SUBAPPLICATION Softkey_Aux_IXA_TO_DataPanel_QXA_BG (* SoftKey ODER AUX auf DataPanel-MI-Ausgang, Hintergrundfarbe SoftKey+AUX Gruen/Weiss, 2 AX-Ausgaenge *)
  (* Standard: 61499-2; Description: Copyright (c) 2026 Meisterschulen am Ostbahnhof This program and the accompanying materials are made available under the terms of the Eclipse Public License 2.0 which is available at https://www.eclipse.org/legal/epl-2.0/ SPDX-License-Identifier: EPL-2.0 *)
  (* Version 1.0, 2026-10-31, Franz Höpfinger, Meisterschulen am Ostbahnhof, Aus Getreidehacke func/Manual/ManFuncTast2 in MyLib::sys verschoben und umbenannt, INIT/INITO/QI/QO ergaenzt, Output und u8SAMember als Parameter. *)
  PACKAGE MyLib::sys;
  IMPORT isobus::UT::Q::const::IDs::ID_NULL;
  IMPORT DataPanel::io::MI::DQ::DataPanel_MI_DO_S;
  IMPORT DataPanel::io::MI::DQ::DataPanel_MI_DO;
  IMPORT DataPanel::io::MI::const::MI;
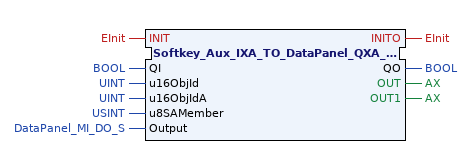
  EVENT_INPUT
    INIT : EInit; (* Initialization Request *)
  END_EVENT
  EVENT_OUTPUT
    INITO : EInit; (* Initialization Confirm *)
  END_EVENT
  VAR_INPUT
    QI : BOOL := TRUE; (* Quality Input - TRUE to enable service *)
    u16ObjId : UINT := ID_NULL; (* Object ID SoftKey *)
    u16ObjIdA : UINT := ID_NULL; (* Object ID AuxFunction2 *)
    u8SAMember : USINT := MI::MI_00; (* DataPanel-MI-Modul (Source Address) *)
    Output : DataPanel::io::MI::DQ::DataPanel_MI_DO_S := DataPanel_MI_DO::Invalid; (* DataPanel-MI-Ausgang *)
  END_VAR
  VAR_OUTPUT
    QO : BOOL; (* Quality Output - TRUE if service executed successfully *)
  END_VAR
  PLUGS
    OUT : adapter::types::unidirectional::AX; (* SoftKey ODER AUX *)
    OUT1 : adapter::types::unidirectional::AX; (* SoftKey ODER AUX (2. Abgriff) *)
  END_PLUGS
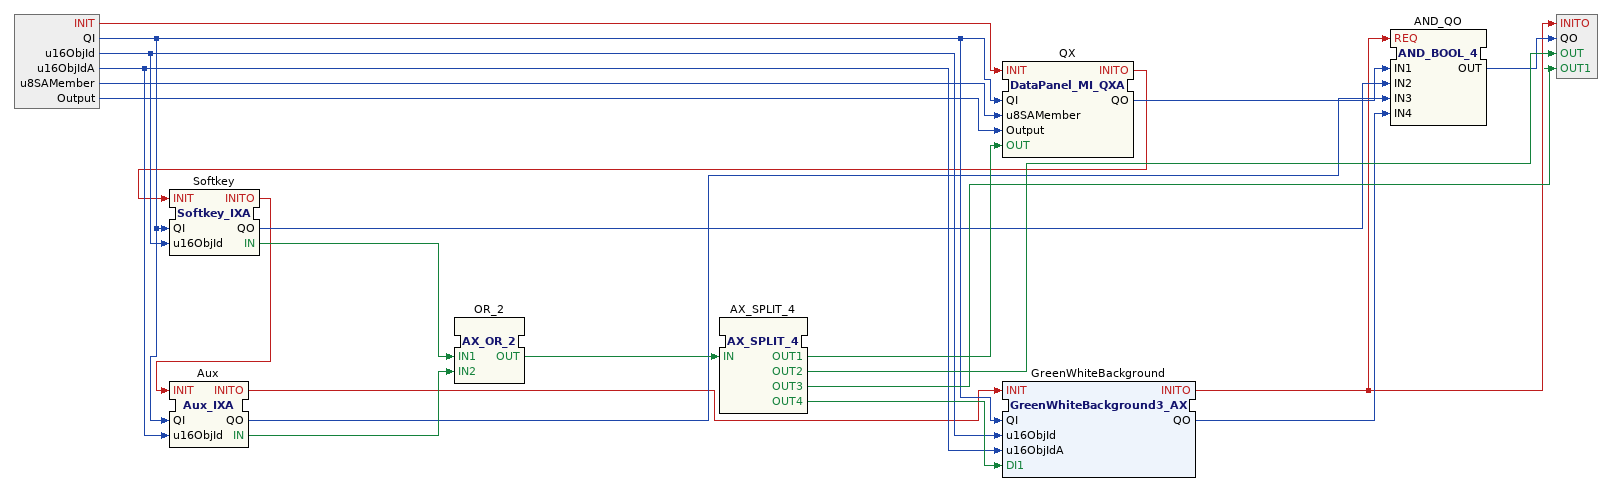
  FBS
    QX : DataPanel::io::MI::DQ::DataPanel_MI_QXA;
    Softkey : isobus::UT::io::Softkey::Softkey_IXA;
    Aux : isobus::UT::io::Auxiliary::IN::Aux_IXA;
    OR_2 : adapter::booleanOperators::AX_OR_2;
    AX_SPLIT_4 : adapter::events::unidirectional::AX_SPLIT_4;
    AND_QO : iec61131::booleanOperators::AND_BOOL_4;
  END_FBS
  SUBAPPS
    GreenWhiteBackground : MyLib::sys::GreenWhiteBackground3_AX;
  END_SUBAPPS
  EVENT_CONNECTIONS
    INIT TO QX.INIT;
    QX.INITO TO Softkey.INIT;
    Softkey.INITO TO Aux.INIT;
    Aux.INITO TO GreenWhiteBackground.INIT;
    GreenWhiteBackground.INITO TO INITO;
    GreenWhiteBackground.INITO TO AND_QO.REQ;
  END_CONNECTIONS
  DATA_CONNECTIONS
    QI TO QX.QI;
    QI TO Softkey.QI;
    QI TO Aux.QI;
    QI TO GreenWhiteBackground.QI;
    u16ObjId TO Softkey.u16ObjId;
    u16ObjIdA TO Aux.u16ObjId;
    u16ObjId TO GreenWhiteBackground.u16ObjId;
    u16ObjIdA TO GreenWhiteBackground.u16ObjIdA;
    u8SAMember TO QX.u8SAMember;
    Output TO QX.Output;
    QX.QO TO AND_QO.IN1;
    Softkey.QO TO AND_QO.IN2;
    Aux.QO TO AND_QO.IN3;
    GreenWhiteBackground.QO TO AND_QO.IN4;
    AND_QO.OUT TO QO;
  END_CONNECTIONS
  ADAPTER_CONNECTIONS
    Softkey.IN TO OR_2.IN1;
    Aux.IN TO OR_2.IN2;
    OR_2.OUT TO AX_SPLIT_4.IN;
    AX_SPLIT_4.OUT1 TO QX.OUT;
    AX_SPLIT_4.OUT2 TO OUT;
    AX_SPLIT_4.OUT3 TO OUT1;
    AX_SPLIT_4.OUT4 TO GreenWhiteBackground.DI1;
  END_CONNECTIONS
END_SUBAPPLICATION
